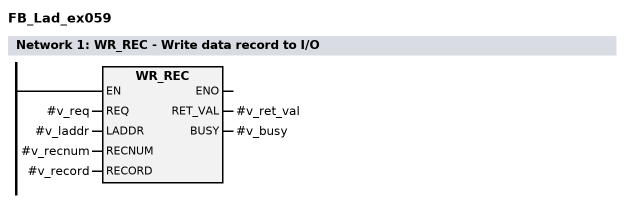
   #v_ret_val := WR_REC(REQ := #v_req,
                        LADDR := #v_laddr,
                        RECNUM := #v_recnum,
                        RECORD := #v_record,
                        BUSY => #v_busy);
END_REGION
END_FUNCTION_BLOCK

FUNCTION_BLOCK "FB_Lad_ex122"   // FB397, LAD
{ S7_Optimized_Access := 'TRUE' }
   VAR_INPUT
      v_operatemode : Byte;
      v_datamode : Byte;
      v_dispclassnr : Array[0..31] of UInt;
      v_lcid : UDInt;
   END_VAR
   VAR_OUTPUT
      v_dataready : Bool;
      v_busy : Bool;
      v_error : Bool;
      v_init : Bool;
      v_status : Word;
   END_VAR
   VAR_IN_OUT
      v_data : AlarmData;
   END_VAR
   VAR
      inst : Get_Alarm;
   END_VAR
BEGIN

REGION Network 1: Get_Alarm - Read pending alarm
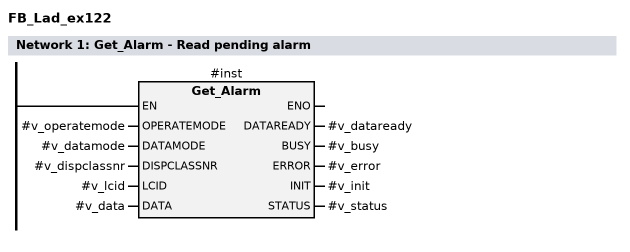
   #inst(OperateMode := #v_operatemode,   // Get_Alarm
         DataMode := #v_datamode,
         DispClassNr := #v_dispclassnr,
         Lcid := #v_lcid,
         Data := #v_data,
         DataReady => #v_dataready,
         Busy => #v_busy,
         Error => #v_error,
         Init => #v_init,
         Status => #v_status);
END_REGION
END_FUNCTION_BLOCK

FUNCTION_BLOCK "FB_Fbd_ex058"   // FB398, FBD
{ S7_Optimized_Access := 'TRUE' }
   VAR_INPUT
      v_req : Bool;
      v_laddr : Hw_Io;
      v_recnum : Byte;
   END_VAR
   VAR_OUTPUT
      v_ret_val : Int;
      v_busy : Bool;
   END_VAR
   VAR_IN_OUT
      v_record : Variant;
   END_VAR
BEGIN

REGION Network 1: RD_REC - Read data record from I/O
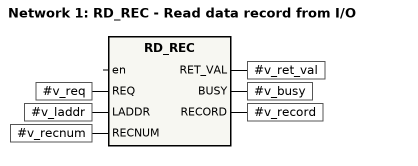
   #v_ret_val := RD_REC(REQ := #v_req,
                        LADDR := #v_laddr,
                        RECNUM := #v_recnum,
                        BUSY => #v_busy,
                        RECORD => #v_record);
END_REGION
END_FUNCTION_BLOCK

FUNCTION_BLOCK "FB_Fbd_ex059"   // FB399, FBD
{ S7_Optimized_Access := 'TRUE' }
   VAR_INPUT
      v_req : Bool;
      v_laddr : Hw_Io;
      v_recnum : Byte;
      v_record : Variant;
   END_VAR
   VAR_OUTPUT
      v_ret_val : Int;
      v_busy : Bool;
   END_VAR
BEGIN

REGION Network 1: WR_REC - Write data record to I/O
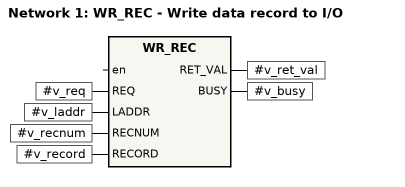
   #v_ret_val := WR_REC(REQ := #v_req,
                        LADDR := #v_laddr,
                        RECNUM := #v_recnum,
                        RECORD := #v_record,
                        BUSY => #v_busy);
END_REGION
END_FUNCTION_BLOCK

FUNCTION_BLOCK "FB_Fbd_ex122"   // FB400, FBD
{ S7_Optimized_Access := 'TRUE' }
   VAR_INPUT
      v_operatemode : Byte;
      v_datamode : Byte;
      v_dispclassnr : Array[0..31] of UInt;
      v_lcid : UDInt;
   END_VAR
   VAR_OUTPUT
      v_dataready : Bool;
      v_busy : Bool;
      v_error : Bool;
      v_init : Bool;
      v_status : Word;
   END_VAR
   VAR_IN_OUT
      v_data : AlarmData;
   END_VAR
   VAR
      inst : Get_Alarm;
   END_VAR
BEGIN

REGION Network 1: Get_Alarm - Read pending alarm
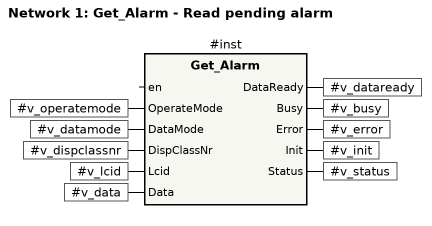
   #inst(OperateMode := #v_operatemode,   // Get_Alarm
         DataMode := #v_datamode,
         DispClassNr := #v_dispclassnr,
         Lcid := #v_lcid,
         Data := #v_data,
         DataReady => #v_dataready,
         Busy => #v_busy,
         Error => #v_error,
         Init => #v_init,
         Status => #v_status);
END_REGION
END_FUNCTION_BLOCK

FUNCTION "FC_SclRt" : Void   // FC1, SCL
{ S7_Optimized_Access := 'TRUE' }
VERSION : 0.1
   VAR_TEMP
      w : Word;
      err : ErrorStruct;
   END_VAR
BEGIN
   // runtime control
           RE_TRIGR();
           #w := GET_ERR_ID();
           GET_ERROR(#err);
           STP();
END_FUNCTION

ORGANIZATION_BLOCK "Main"   // OB1, LAD, ProgramCycle
TITLE = "Main Program Sweep (Cycle)"
{ S7_Optimized_Access := 'TRUE' }
VERSION : 0.1
   VAR_INPUT
      Initial_Call : Bool;   // Initial call of this OB
      Remanence : Bool;   // =True, if remanent data are available
   END_VAR
BEGIN
END_ORGANIZATION_BLOCK